Fanuc KAREL source: KA00126.KL

PROGRAM KA00126
%NOLOCKGROUP
VAR
  SRC: ARRAY[2] OF BYTE
  DST: XYZWPR
BEGIN
  SRC[1] = 2
  DST = SRC[1]
END KA00126
